(* Test host that nests an FB_ATM, the way a device FB would. Its references are
   bound in its own FB_Init, which runs after the nested FB_ATM was constructed
   from them, so the nested FB_ATM first sees nil references. CallAfterInit
   re-supplies them through fbATM.CallAfterInitATM. *)
{attribute 'call_after_init'}
FUNCTION_BLOCK FB_ATMHost
VAR
    {attribute 'no_copy'}
    aiMotionStage         : REFERENCE TO ARRAY[1..MotionConstants.MAX_STATE_MOTORS] OF I_MotionStage;
    {attribute 'no_copy'}
    astPositionState      : REFERENCE TO ARRAY[1..MotionConstants.MAX_STATE_MOTORS]
                                            OF ARRAY[1..GeneralConstants.MAX_STATES] OF ST_PositionState;
    {attribute 'no_copy'}
    fbFFHWO               : REFERENCE TO FB_HardwareFFOutput;
    {attribute 'no_copy'}
    fbArbiter             : REFERENCE TO FB_Arbiter;
    sDeviceName           : STRING;
    sTransitionKey        : STRING;
    bEnableBeamParams     : BOOL;
    bEnablePositionLimits : BOOL;
    bReadDBNow            : BOOL;
    {attribute 'no_copy'}
    bFileReaderBusy       : REFERENCE TO BOOL;
    {attribute 'no_copy'}
    bFileReaderError      : REFERENCE TO BOOL;

    fbATM : FB_ATM(
        aiMotionStage         := aiMotionStage,
        astPositionState      := astPositionState,
        fbFFHWO               := fbFFHWO,
        fbArbiter             := fbArbiter,
        sDeviceName           := sDeviceName,
        sTransitionKey        := sTransitionKey,
        bEnableBeamParams     := bEnableBeamParams,
        bEnablePositionLimits := bEnablePositionLimits,
        bReadDBNow            := bReadDBNow,
        bFileReaderBusy       := bFileReaderBusy,
        bFileReaderError      := bFileReaderError
    );
END_VAR

fbATM();

(* The nested fbATM ran its own CallAfterInit before this one, with nil
   references. Re-supplies them and redoes its wiring. *)
{attribute 'call_after_init'}
METHOD CallAfterInit
fbATM.CallAfterInitATM(
    aiMotionStage         := aiMotionStage,
    astPositionState      := astPositionState,
    fbFFHWO               := fbFFHWO,
    fbArbiter             := fbArbiter,
    sDeviceName           := sDeviceName,
    sTransitionKey        := sTransitionKey,
    bEnableBeamParams     := bEnableBeamParams,
    bEnablePositionLimits := bEnablePositionLimits,
    bReadDBNow            := bReadDBNow,
    bFileReaderBusy       := bFileReaderBusy,
    bFileReaderError      := bFileReaderError
);
END_METHOD

(* Stores the injected references and values in this FB's fields. *)
{attribute 'analysis' := '-33'}
METHOD FB_Init : BOOL
VAR_INPUT
    bInitRetains           : BOOL;
    bInCopyCode            : BOOL;
    aiMotionStage          : REFERENCE TO ARRAY[1..MotionConstants.MAX_STATE_MOTORS] OF I_MotionStage;
    astPositionState       : REFERENCE TO ARRAY[1..MotionConstants.MAX_STATE_MOTORS]
                                            OF ARRAY[1..GeneralConstants.MAX_STATES] OF ST_PositionState;
    fbFFHWO                : REFERENCE TO FB_HardwareFFOutput;
    fbArbiter              : REFERENCE TO FB_Arbiter;
    sDeviceName            : STRING;
    sTransitionKey         : STRING;
    bEnableBeamParams      : BOOL;
    bEnablePositionLimits  : BOOL;
    bReadDBNow             : BOOL;
    bFileReaderBusy        : REFERENCE TO BOOL;
    bFileReaderError       : REFERENCE TO BOOL;
END_VAR
THIS^.aiMotionStage         REF= aiMotionStage;
THIS^.astPositionState      REF= astPositionState;
THIS^.fbFFHWO               REF= fbFFHWO;
THIS^.fbArbiter             REF= fbArbiter;
THIS^.sDeviceName           := sDeviceName;
THIS^.sTransitionKey        := sTransitionKey;
THIS^.bEnableBeamParams     := bEnableBeamParams;
THIS^.bEnablePositionLimits := bEnablePositionLimits;
THIS^.bReadDBNow            := bReadDBNow;
THIS^.bFileReaderBusy       REF= bFileReaderBusy;
THIS^.bFileReaderError      REF= bFileReaderError;
END_METHOD

END_FUNCTION_BLOCK

(* stored: Version 1.1.0.1
   POU FB_ATMHost: Id {0bbfe163-a749-433e-a69a-6c897167c9b3}, SpecialFunc None
   Method CallAfterInit: Id {69049f69-7b85-471f-984b-eb2e5edfc54d}
   Method FB_Init: Id {5f37f847-f7db-4c88-a1bc-b7b0b1b9f132} *)
